FUNCTION_BLOCK FTS_MCMoveVelocity
VAR_IN_OUT
	stAxis: ST_Axis;
END_VAR
VAR_INPUT
	bExecute: BOOL;
	bCollsionNotValid: BOOL := FALSE;
	fVelocity: LREAL;
	fAcceleration: LREAL;
	fDeceleration: LREAL;
	fJerk: LREAL;
	fGap: LREAL;
	eDirection: E_Direction;
	eBufferMode: E_MCBufferMode := E_MCBufferMode.ABORTING;
END_VAR
VAR_OUTPUT
	bInVelocity: BOOL;
	bActive: BOOL;
	bBusy: BOOL;
	bCommandAborted: BOOL;
	bError: BOOL;
	nErrorID: UDINT;
END_VAR
VAR
	_bNcStart: BOOL;
	_bSegDone: BOOL;
	_bPathCalDone: BOOL := FALSE;
	_bParamError: BOOL := FALSE;
	_bCollisionChecked: BOOL;
	_nStep: INT;
	_nSysType: UINT;
	_nCycleCount: UDINT := 0;
	///02.24
	_nLastNcCycleCounter: UDINT;
	///02.24
	_nDealtNcCycleCounter: UDINT;
	///02.24
	_nLastCycleCounter: UDINT;
	///02.24
	_nDealtCycleCounter: UDINT;
	_fPostion: LREAL;
	_fDec: LREAL;
	_fDistance: LREAL;
	_fGap: LREAL;
	_fClampLength: LREAL;
	_fAcc: LREAL;
	_fPrePosition: LREAL;
	_fPrePositionTemp: LREAL;
	_fSetVelo: LREAL;
	_eCommand: E_Command;
	_pPremover: POINTER TO ST_Axis;
	_stTimeInfo: ST_TimeRef;
	_stPathRef: ST_PathRef;
	_stNoPathRef: ST_PathRef;
	_stAxisNo: ST_Axis;
	_fbTrig: R_TRIG;
	///03.04
	_fbEnbleTrig: F_TRIG;
	_fbDoneTon: TON;
	_fbWaitTon: TON;
	_fbTraPlanning: FB_TrajectoryPlanning;
END_VAR
VAR CONSTANT
	//fNcCycle: REAL := 0.001;
	tcDoneTime: TIME := TIME#100ms;
	//tcWaitTime: TIME := TIME#500ms;
	//tcCalcuTime: TIME := TIME#33m20s0ms;
	fPositivePosSet: LREAL := 500000000;
	fNegativePosSet: LREAL := -500000000;
	//fGapSet: LREAL := 100000;
END_VAR


IF (eDirection=E_Direction.DIRECTION_POSITIVE)THEN
	IF (stAxis.stAxisStatus.pPremover=0)THEN 
		_pPremover:=ADR(_stAxisNo);
	ELSE
		_pPremover:=stAxis.stAxisStatus.pPremover;
	END_IF
ELSE
	IF (stAxis.stAxisStatus.pAftermover=0)THEN 
		_pPremover:=ADR(_stAxisNo);
	ELSE
		_pPremover:=stAxis.stAxisStatus.pAftermover;
	END_IF

END_IF
A_CommandCheck();

// 02.24增加task事件判断
IF (_nStep<>0)THEN 
	_nCycleCount:=_nCycleCount+1;
ELSE
	_nCycleCount:=0;
END_IF


CASE _nStep OF 
	0:
	    
	    IF NOT bExecute THEN 
		   bError:=FALSE;
		   nErrorId:=0;
		   bInVelocity:=FALSE;
		   bCommandAborted:=FALSE;
		  
		   _eCommand:=E_Command.COMMAND_IDLE;
	   END_IF   
	   RETURN;
	10:
	    bBusy:=TRUE;
	    bError:=FALSE;
	    bCommandAborted:=FALSE;
	    nErrorID:=0;
		bActive:=FALSE;
		bInVelocity:=FALSE;
		 A_ParamCheck();
		 IF (stAxis.stPLCTONC.eCommand<>E_Command.COMMAND_MOVEVELOCITY)THEN
			 IF NOT stAxis.stPLCTONC.bNcStart THEN
				 _nStep:= 20;
			 END_IF
		 ELSE
			 stAxis.stPLCTONC.bNcStart:=FALSE;
		     _nStep:= 20;
		 END_IF
		 //stAxis.stPLCTONC.bNcStart:=FALSE;
        //_nStep:=10+_nStep;
		
	    IF _bParamError  THEN 
			 _nStep:= 100;
			 _bParamError:=FALSE;
		END_IF
		
	20:  //calculate path 
	    bActive:=TRUE;
	    A_CalcutaPath();
     
		stAxis.stAxisStatus.bContinuousMotion:=TRUE;
		stAxis.stAxisStatus.bDiscreteMotion:=FALSE;
		stAxis.stAxisStatus.bSynchronizedMotion:=FALSE;
		stAxis.stPLCTONC.eCommand:=E_Command.COMMAND_MOVEVELOCITY;
		_eCommand:=stAxis.stPLCTONC.eCommand;
		_bCollisionChecked:=FALSE;
		IF _bPathCalDone THEN
			stAxis.stPLCTONC.bNcEnable:=TRUE;
		    stAxis.stPLCTONC.bNcStart:=TRUE;
		    //stAxis.stPLCTONC.eCommand:=E_Command.COMMAND_MOVEVELOCITY;
			// _eCommand:=stAxis.stPLCTONC.eCommand;
			stAxis.stPLCTONC.ePlanningMode:=E_PlanningMode.PLANNINGMODE_TSHAPED;
		    stAxis.stAxisStatus.bConstantVelocity:=TRUE;
	
			_nStep:=25;
			_bPathCalDone:=FALSE;
		END_IF
		IF _bSegDone THEN 
			_nStep:=0;
			 bBusy:=FALSE;
	         bActive:=FALSE;
			 bInVelocity:=TRUE;
			 _bSegDone:=FALSE;
			 _bCollisionChecked:=TRUE;
			 stAxis.stPLCTONC.eCommand:=E_Command.COMMAND_IDLE;
			_eCommand:=E_Command.COMMAND_IDLE;
			
		END_IF
	25:
	    _nStep:=30;
		// stAxis.stPLCTONC.bNcStart:=FALSE;
		  //自动计算nc task和规划task 02.24
		 _nDealtCycleCounter:=_nCycleCount-_nLastCycleCounter;
		 _nDealtNcCycleCounter:=stAxis.stAxisStatus.nNcCycleCounter_WP-_nLastNcCycleCounter;
		 IF (_nDealtCycleCounter< _nDealtNcCycleCounter)THEN
			  stAxis.stPLCTONC.bNcStart:=FALSE;     //12.27
		 END_IF
    30:
         stAxis.stPLCTONC.bNcStart:=FALSE;
		 
	     IF (stAxis.stPLCTONC.stStartPosition.fVelocity<stAxis.stPLCTONC.fTargetVelocity )THEN
              IF (stAxis.stNcTOPLC.fActVelo>=_fSetVelo)THEN 
		              bInVelocity:=TRUE;
			  END_IF
		 ELSE
			  IF (stAxis.stNcTOPLC.fActVelo<=_fSetVelo)THEN 
		              bInVelocity:=TRUE;
			  END_IF
	     END_IF
		 IF (stAxis.stNcTOPLC.nAxisState=2)THEN
			   _nStep:=0; 
			  
			   bCommandAborted:=FALSE;
			   bBusy:=FALSE;
			   bActive:=FALSE;
			   bInVelocity:=FALSE;
			   stAxis.stAxisStatus.bConstantVelocity:=FALSE;
			  
			   stAxis.stAxisStatus.bContinuousMotion:=FALSE;
			   stAxis.stPLCTONC.eCommand:=E_Command.COMMAND_IDLE;
			   _eCommand:=E_Command.COMMAND_IDLE;
			   stAxis.stPLCTONC.ePlanningMode:=E_PlanningMode.PLANNINGMODE_NONE;
			   stAxis.stPLCTONC.bNcStart:=FALSE;
			   stAxis.stPLCTONC.bNcEnable:=FALSE;
			   _bCollisionChecked:=TRUE;
	    END_IF
       
    
    //  disEnable     
    40:
	    IF (stAxis.stAxisStatus.nNcCycleCounter<>0)THEN
			A_StopPathGeneration();
			 stAxis.stPLCTONC.bNcStart:=TRUE;
			_nStep:=_nStep+10;
	    ELSE
		  (* _nStep:=0;
           bInVelocity:=FALSE;
		   bCommandAborted:=TRUE;
		   bBusy:=FALSE;
		   bActive:=FALSE;
		   stAxis.stAxisStatus.bMoving:=FALSE;
		   stAxis.stPLCTONC.bNcStart:=FALSE; 
		   stAxis.stAxisStatus.bConstantVelocity:=FALSE;
	       stAxis.stAxisStatus.bContinuousMotion:=FALSE;
		   _bCollisionChecked:=FALSE;
		   stAxis.stPLCTONC.ePlanningMode:=E_PlanningMode.PLANNINGMODE_NONE;
		   stAxis.stPLCTONC.eCommand:=E_Command.COMMAND_IDLE;
		   _eCommand:=E_Command.COMMAND_IDLE;*)
		   _nStep:=60;
		END_IF 
	   
    50:
	    IF (stAxis.stNcTOPLC.nAxisState=2)THEN
	       _nStep:=_nStep+10; 
		   stAxis.stPLCTONC.bNcStart:=FALSE;
           _fbDoneTon(IN:=FALSE, PT:=tcDoneTime , Q=> , ET=> );
	   
        END_IF
	60:
    	
	   // _fbDoneTon(IN:=TRUE, PT:=tcDoneTime , Q=> , ET=> );
       // IF _fbDoneTon.Q THEN
			
			 _fbDoneTon(IN:=FALSE, PT:=tcDoneTime , Q=> , ET=> );
			  _nStep:=0;
			   bCommandAborted:=TRUE;
			   bInVelocity:=FALSE;
		       bBusy:=FALSE;
		       bActive:=FALSE;
			  stAxis.stAxisStatus.bContinuousMotion:=FALSE;
			  stAxis.stAxisStatus.bConstantVelocity:=FALSE;
			  stAxis.stPLCTONC.bNcEnable:=FALSE;
			  stAxis.stPLCTONC.ePlanningMode:=E_PlanningMode.PLANNINGMODE_NONE;
			  stAxis.stPLCTONC.eCommand:=E_Command.COMMAND_IDLE;
			  _eCommand:=E_Command.COMMAND_IDLE;
			  _bCollisionChecked:=FALSE;
	    // END_IF	 
		
    100: (************error handle***********)
         bBusy:=FALSE;
	     bError:=TRUE;
	     bInVelocity:=FALSE;
		 bActive:=FALSE;
	     bCommandAborted:=FALSE;
	     stAxis.stAxisStatus.bError:=TRUE;
		 stAxis.stAxisStatus.nErrorId:=nErrorId;
	     _nStep:=0;
		 stAxis.stPLCTONC.bNcStart:=FALSE;
		 stAxis.stPLCTONC.bNcEnable:=FALSE;
		 stAxis.stAxisStatus.bConstantVelocity:=FALSE;
		 stAxis.stPLCTONC.ePlanningMode:=E_PlanningMode.PLANNINGMODE_NONE;
	     stAxis.stPLCTONC.eCommand:=E_Command.COMMAND_IDLE;
	
		 stAxis.stAxisStatus.bConstantVelocity:=FALSE;
		 stAxis.stAxisStatus.bContinuousMotion:=FALSE;
		 _bCollisionChecked:=FALSE;
		 
	110:
	     bCommandAborted:=TRUE;
	     bBusy:=FALSE;
	     bInVelocity:=FALSE;
	     bActive:=FALSE;
	     _nStep:=0; 
	     stAxis.stAxisStatus.bConstantVelocity:=FALSE;
	     //stAxis.stAxisStatus.bContinuousMotion:=FALSE;
	     _bCollisionChecked:=FALSE;
END_CASE


A_UpstateStatus();

ACTION A_CalcutaPath:


stAxis.stPLCTONC.stStartPosition.fPosition:=stAxis.stNcTOPLC.fActPos;
stAxis.stPLCTONC.stStartPosition.fVelocity:=stAxis.stNcTOPLC.fActVelo;
stAxis.stPLCTONC.stStartPosition.fAccleration:=fAcceleration;
stAxis.stPLCTONC.stStartPosition.fDeceleration:=fDeceleration;
stAxis.stPLCTONC.stStartPosition.fbJerk:=fJerk;

stAxis.stPLCTONC.fTargetVelocity:=_fSetVelo;
stAxis.stPLCTONC.fSetVelocity:=_fSetVelo;  //04.25
stAxis.stPLCTONC.stEndPosition.fVelocity:=0;
stAxis.stPLCTONC.stEndPosition.fAccleration:=_fAcc;
stAxis.stPLCTONC.stEndPosition.fDeceleration:=_fDec;
stAxis.stPLCTONC.stEndPosition.fbJerk:=fJerk;
IF(eDirection=E_Direction.DIRECTION_POSITIVE)THEN 
	stAxis.stPLCTONC.stEndPosition.fPosition:=fPositivePosSet+stAxis.stPLCTONC.stStartPosition.fPosition;
ELSE
   stAxis.stPLCTONC.stEndPosition.fPosition:=fNegativePosSet+stAxis.stPLCTONC.stStartPosition.fPosition;
END_IF

stAxis.stPLCTONC.nSysType:=_nSysType;
IF (_nSysType=1)OR (_nSysType=4) THEN 
	stAxis.stPLCTONC.nSysType:=2;
END_IF
//stAxis.stAxisStatus.stPathRef.fGap:=_fGap;
//stAxis.stAxisStatus.stPathRef.fGap:=0;
stAxis.stAxisStatus.stPathRef.fGap:=_fClampLength;
stAxis.stAxisStatus.stPathRef.fSetGap:=_fGap;

IF (_pPremover^.stNcTOPLC.nAxisId<>0)AND NOT bCollsionNotValid THEN
	IF(eDirection=E_Direction.DIRECTION_POSITIVE)THEN 
	    IF _pPremover^.stAxisStatus.bPositiveDirection THEN 
			_fPrePosition:=FC_FindPosition(pPathData:=_pPremover^.stAxisStatus.stPathRef.aSafePath )-_fGap;
			IF (_pPremover^.stNcTOPLC.fActPos<stAxis.stNcTOPLC.fActPos)AND(_nSysType=3)THEN    //cycle positive move
				_fPrePosition:=_fPrePosition+stAxis.stNcTOPLC.fModuloFactor;
			END_IF 
			
		ELSE
			_fPrePosition:=FC_FindPosition(pPathData:=_pPremover^.stAxisStatus.stPathRef.aExecutablePath)-_pPremover^.stAxisParam.fClampLength*0.5-_fGap;
			IF (_pPremover^.stNcTOPLC.fActPos<stAxis.stNcTOPLC.fActPos)AND(_nSysType=3)THEN    //cycle positive move
				_fPrePosition:=_fPrePosition+stAxis.stNcTOPLC.fModuloFactor;
			END_IF 
			
		END_IF
		_fPrePositionTemp:=_fPrePosition;
		IF (_pPremover^.stAxisStatus.nNcCycleCounter=0)THEN 
			 IF (_pPremover^.stNcTOPLC.fActPos<stAxis.stNcTOPLC.fActPos)THEN    //cycle positive move
					 _fPrePosition:=_pPremover^.stNcTOPLC.fActPos+stAxis.stNcTOPLC.fModuloFactor-_pPremover^.stAxisParam.fClampLength*0.5-_fClampLength-ABS(fGap);
			 ELSE
					 _fPrePosition:=_pPremover^.stNcTOPLC.fActPos--_pPremover^.stAxisParam.fClampLength*0.5-_fClampLength-ABS(fGap);
			 END_IF 
		END_IF
		IF (_fPrePosition<stAxis.stNcTOPLC.fActPos)THEN 
			   _bSegDone:=TRUE;
               RETURN; 
		 END_IF
		 IF (stAxis.stPLCTONC.stEndPosition.fPosition>_fPrePosition)THEN
			stAxis.stPLCTONC.stEndPosition.fPosition:=_fPrePosition;
		 END_IF
		 
    ELSE
	     IF _pPremover^.stAxisStatus.bNegativeDirection THEN // 负向
			_fPrePosition:=FC_FindPosition(pPathData:=_pPremover^.stAxisStatus.stPathRef.aSafePath )+_fGap;
			IF (_pPremover^.stNcTOPLC.fActPos>stAxis.stNcTOPLC.fActPos)AND(_nSysType=3)THEN    //cycle negative  move
				_fPrePosition:=_fPrePosition-stAxis.stNcTOPLC.fModuloFactor;
				 
			END_IF
		ELSE
			_fPrePosition:=FC_FindPosition(pPathData:=_pPremover^.stAxisStatus.stPathRef.aExecutablePath )+_pPremover^.stAxisParam.fClampLength*0.5+_fGap;
			IF (_pPremover^.stNcTOPLC.fActPos>stAxis.stNcTOPLC.fActPos)AND(_nSysType=3)THEN    //cycle negative  move
				_fPrePosition:=_fPrePosition-stAxis.stNcTOPLC.fModuloFactor;
			END_IF
		END_IF
		_fPrePositionTemp:=_fPrePosition;
		IF (_pPremover^.stAxisStatus.nNcCycleCounter=0)THEN
			 IF (_pPremover^.stNcTOPLC.fActPos>stAxis.stNcTOPLC.fActPos)THEN    //cycle positive move
					 
					 _fPrePosition:=_pPremover^.stNcTOPLC.fActPos-stAxis.stNcTOPLC.fModuloFactor+_pPremover^.stAxisParam.fClampLength*0.5+_fClampLength+ABS(fGap);
			 ELSE
					 _fPrePosition:=_pPremover^.stNcTOPLC.fActPos+_pPremover^.stAxisParam.fClampLength*0.5+_fClampLength+ABS(fGap);
			 END_IF
		 END_IF
		 IF (_fPrePosition>stAxis.stNcTOPLC.fActPos)THEN 
			   _bSegDone:=TRUE;
               RETURN; 
		 END_IF
		 IF (stAxis.stPLCTONC.stEndPosition.fPosition<_fPrePosition)THEN
			stAxis.stPLCTONC.stEndPosition.fPosition:=_fPrePosition;
		 END_IF
    END_IF 
  
END_IF
_fDistance:=ABS(stAxis.stPLCTONC.stEndPosition.fPosition-stAxis.stPLCTONC.stStartPosition.fPosition);
	
IF (_fDistance<=0)THEN 
   _bSegDone:=TRUE;
	 RETURN ;
END_IF

IF (eDirection=E_Direction.DIRECTION_POSITIVE)THEN
	stAxis.stAxisStatus.bPositiveDirection:=TRUE;
	stAxis.stAxisStatus.bNegativeDirection:=FALSE;
ELSE
    stAxis.stAxisStatus.bPositiveDirection:=FALSE;
	stAxis.stAxisStatus.bNegativeDirection:=TRUE;
END_IF 
_bPathCalDone:=TRUE;
END_ACTION

ACTION A_CommandCheck:

//注意优先级，最下面优先级最高

_fbTrig(CLK:=bExecute , Q=> );
IF _fbTrig.Q  THEN
	IF (NOT stAxis.stAxisStatus.bEnabled) OR stAxis.stAxisStatus.bError OR stAxis.stAxisStatus.bStopping THEN 
		_nStep:=100;
		//bError:=TRUE;
		nErrorID:=29703;
		RETURN;
	END_IF
	
	_nStep:=10;
END_IF

//command aborted   /12/1
IF (stAxis.stPLCTONC.eCommand<>E_Command.COMMAND_MOVEVELOCITY) AND (_nStep<>0)AND(_eCommand=E_Command.COMMAND_MOVEVELOCITY)THEN 
	_nStep:=110; 
END_IF

// disEnable
_fbEnbleTrig(CLK:=stAxis.stAxisStatus.bEnabled, Q=> );
IF _fbEnbleTrig.Q THEN 
	//bCommandAborted:=TRUE;
	IF (_nStep=0)THEN
		bBusy:=FALSE;
	    bInVelocity:=FALSE;
	    bActive:=FALSE;
	    _nStep:=0; 
		 _bCollisionChecked:=FALSE;
	ELSE
		//_nStep:=40;   //规划
		_nStep:=60;     //不规划
	END_IF
	
END_IF
END_ACTION

ACTION A_Init:
_bPathCalDone:=FALSE;
_stPathRef:=_stNoPathRef;
bCommandAborted:=FALSE;
 _bSegDone:=false;
END_ACTION

ACTION A_MeasureIn:

_fClampLength:=stAxis.stAxisParam.fClampLength*0.5;

IF ABS(fVelocity)>stAxis.stAxisParam.stDynamicDefault.fMaxVelocity THEN 
	_fSetVelo:= stAxis.stAxisParam.stDynamicDefault.fMaxVelocity ;
ELSE
	_fSetVelo:= ABS(fVelocity) ;
END_IF

IF (fGap<>0)THEN 
   _fGap :=_fClampLength+ABS(fGap);
     
ELSE
  _fGap :=_fClampLength+ABS(stAxis.stAxisParam.fGap);
 
END_IF

IF (fAcceleration=0) THEN 
	_fAcc:=stAxis.stAxisParam.stDynamicDefault.fDefaultAccelaration;
ELSE
	_fAcc:=ABS(fAcceleration);
	IF (fAcceleration>stAxis.stAxisParam.stDynamicDefault.fMaxAccelaration)THEN
		_fAcc:=stAxis.stAxisParam.stDynamicDefault.fMaxAccelaration;
	END_IF
END_IF


IF (fDeceleration=0) THEN
   _fDec:=stAxis.stAxisParam.stDynamicDefault.fDefaultDeceleration;
ELSE 
	_fDec:=ABS(fDeceleration);
	IF (fDeceleration>stAxis.stAxisParam.stDynamicDefault.fMaxDeceleration)THEN
		_fDec:=stAxis.stAxisParam.stDynamicDefault.fMaxDeceleration;
	END_IF
END_IF

IF (_fAcc<>_fDec)THEN
	_fDec:=_fAcc;
END_IF

_nSysType:=stAxis.stAxisParam.stRoadParam.nSysType;
END_ACTION

ACTION A_ParamCheck:
A_MeasureIn();

IF(fVelocity=0) THEN       // param error 
	_bParamError:=TRUE;
	nErrorID:=29708;
	RETURN;
END_IF
END_ACTION

ACTION A_StopPathGeneration:
_fPostion:=0.5*stAxis.stNcTOPLC.fActVelo*stAxis.stNcTOPLC.fActVelo/_fDec;
//_fPostion:=0.5*stAxis.stNcTOPLC.fActVelo*stAxis.stNcTOPLC.fActVelo/stAxis.stAxisParam.stDynamicDefault.fMaxDeceleration;
IF stAxis.stAxisStatus.bPositiveDirection THEN
	 stAxis.stPLCTONC.stEndPosition.fPosition:=_fPostion+stAxis.stNcTOPLC.fActPos;
ELSE
	stAxis.stPLCTONC.stEndPosition.fPosition:=stAxis.stNcTOPLC.fActPos-_fPostion;
END_IF

stAxis.stPLCTONC.fTargetVelocity:=stAxis.stNcTOPLC.fActVelo;
stAxis.stPLCTONC.stEndPosition.fVelocity:=0;
stAxis.stPLCTONC.stEndPosition.fAccleration:=_fDec;
stAxis.stPLCTONC.stEndPosition.fDeceleration:=_fDec;
END_ACTION

ACTION A_UpstateStatus:
//stAxis.stAxisStatus.nCollState.3:=_bCollisionChecked;;
stAxis.stAxisStatus.bCollisionStoped:=_bCollisionChecked;

//02.24
_nLastCycleCounter:=_nCycleCount;
_nLastNcCycleCounter:=stAxis.stAxisStatus.nNcCycleCounter_WP;
END_ACTION

END_FUNCTION_BLOCK

(* stored: Version 1.1.0.1, ProductVersion 3.1.4024.12
   POU FTS_MCMoveVelocity: Id {aef16a97-36a6-4538-928f-1ab8bacdcc3e}, SpecialFunc None
   Action A_CalcutaPath: Id {8ba50a66-3e7a-48a9-b684-8ac2677645ab}
   Action A_CommandCheck: Id {2788fcbd-313a-4838-a366-0c14e0752498}
   Action A_Init: Id {c94b88cc-3ea0-4b12-bdb5-130f5467b173}
   Action A_MeasureIn: Id {72c1fc1c-17f9-49e4-b664-328b4d42d501}
   Action A_ParamCheck: Id {9260b475-9ce5-45a5-8862-53f5989bdb33}
   Action A_StopPathGeneration: Id {e0eb3274-7b98-484f-8c69-20f2dcbbbef7}
   Action A_UpstateStatus: Id {36a5f609-6901-4995-95de-2d4d922aba1e} *)
